// TIA Portal V19 export
TYPE "VFD"
   STRUCT
      STW : Word;   // CONTROL WORD
      ZSW : Word;   // STATUS WORD
      HIW : Word;   // ACTUAL SPEED
      HSW : Word;   // SPEED SETPOINT
      ADDR : UInt := 1;   // ADDRESS
      FAULT : Bool;
      "LOCAL/REMOTE" : Int;
   END_STRUCT;
END_TYPE
